(* IEC 61131-3 sources: trust-platform/examples/OSCAT/booster_commissioning_decorator/oop/src, 3 files *)

(* ---- Main.st ---- *)
(* Pattern role: ISignalSource is the contract boundary for the Decorator example. *)
INTERFACE ISignalSource
    PROPERTY Value : REAL
    GET
    END_GET
    END_PROPERTY

    PROPERTY Quality : BYTE
    GET
    END_GET
    END_PROPERTY

    METHOD Update
    END_METHOD
END_INTERFACE

(* Pattern role: IPump is the contract boundary for the Decorator example. *)
INTERFACE IPump
    PROPERTY IsRunning : BOOL
    GET
    END_GET
    END_PROPERTY

    METHOD Run
    VAR_INPUT
        SpeedReference : REAL;
    END_VAR
    END_METHOD

    METHOD Stop
    END_METHOD
END_INTERFACE

(* Pattern role: RealPressureSource is a concrete implementation in the Decorator example. *)
FUNCTION_BLOCK RealPressureSource IMPLEMENTS ISignalSource
VAR
    ValueValue : REAL;
    QualityValue : BYTE := BYTE#2;
END_VAR

METHOD PUBLIC Configure
VAR_INPUT
    PressureBar : REAL;
    QualityCode : BYTE;
END_VAR
ValueValue := PressureBar;
QualityValue := QualityCode;
END_METHOD

METHOD PUBLIC Update
END_METHOD

PUBLIC PROPERTY Value : REAL
GET
    Value := ValueValue;
END_GET
END_PROPERTY

PUBLIC PROPERTY Quality : BYTE
GET
    Quality := QualityValue;
END_GET
END_PROPERTY
END_FUNCTION_BLOCK

(* Pattern role: SimulatedPressureDecorator is a concrete implementation in the Decorator example. *)
FUNCTION_BLOCK SimulatedPressureDecorator IMPLEMENTS ISignalSource
VAR
    RealSourceRef : ISignalSource;
    SineGen : SineSignalGenerator;
    UseSimulationValue : BOOL;
    ValueValue : REAL;
    QualityValue : BYTE;
END_VAR

METHOD PUBLIC Wrap
VAR_INPUT
    RealSource : ISignalSource;
    UseSimulation : BOOL;
END_VAR
RealSourceRef := RealSource;
UseSimulationValue := UseSimulation;
SineGen.Initialize();
SineGen.Configure(Period := T#10s, Amplitude := REAL#0.5, Offset := REAL#4.5, Delay := REAL#0.0);
END_METHOD

METHOD PUBLIC SetSimulation
VAR_INPUT
    Enabled : BOOL;
END_VAR
UseSimulationValue := Enabled;
END_METHOD

METHOD PUBLIC Update
RealSourceRef.Update();
IF UseSimulationValue THEN
    ValueValue := SineGen.Update();
    QualityValue := BYTE#2;
ELSE
    ValueValue := RealSourceRef.Value;
    QualityValue := RealSourceRef.Quality;
END_IF;
END_METHOD

PUBLIC PROPERTY Value : REAL
GET
    Value := ValueValue;
END_GET
END_PROPERTY

PUBLIC PROPERTY Quality : BYTE
GET
    Quality := QualityValue;
END_GET
END_PROPERTY

PUBLIC PROPERTY UsingSimulation : BOOL
GET
    UsingSimulation := UseSimulationValue;
END_GET
END_PROPERTY
END_FUNCTION_BLOCK

(* Pattern role: RealPumpDrive is a concrete implementation in the Decorator example. *)
FUNCTION_BLOCK RealPumpDrive IMPLEMENTS IPump
VAR
    RunningValue : BOOL;
    LastSpeedValue : REAL;
END_VAR

METHOD PUBLIC Run
VAR_INPUT
    SpeedReference : REAL;
END_VAR
LastSpeedValue := SpeedReference;
RunningValue := SpeedReference > REAL#0.0;
END_METHOD

METHOD PUBLIC Stop
LastSpeedValue := REAL#0.0;
RunningValue := FALSE;
END_METHOD

PUBLIC PROPERTY IsRunning : BOOL
GET
    IsRunning := RunningValue;
END_GET
END_PROPERTY

PUBLIC PROPERTY LastSpeed : REAL
GET
    LastSpeed := LastSpeedValue;
END_GET
END_PROPERTY
END_FUNCTION_BLOCK

(* Pattern role: CommissioningOutputDriver is a concrete implementation in the Decorator example. *)
FUNCTION_BLOCK CommissioningOutputDriver IMPLEMENTS IPump
VAR
    RealPump : IPump;
    LoopbackOnlyValue : BOOL;
    LastCommandedSpeedValue : REAL;
END_VAR

METHOD PUBLIC Wrap
VAR_INPUT
    Pump : IPump;
    LoopbackOnly : BOOL;
END_VAR
RealPump := Pump;
LoopbackOnlyValue := LoopbackOnly;
END_METHOD

METHOD PUBLIC SetLoopback
VAR_INPUT
    Enabled : BOOL;
END_VAR
LoopbackOnlyValue := Enabled;
END_METHOD

METHOD PUBLIC Run
VAR_INPUT
    SpeedReference : REAL;
END_VAR
LastCommandedSpeedValue := SpeedReference;
IF NOT LoopbackOnlyValue THEN
    RealPump.Run(SpeedReference := SpeedReference);
END_IF;
END_METHOD

METHOD PUBLIC Stop
LastCommandedSpeedValue := REAL#0.0;
IF NOT LoopbackOnlyValue THEN
    RealPump.Stop();
END_IF;
END_METHOD

PUBLIC PROPERTY IsRunning : BOOL
GET
    IF LoopbackOnlyValue THEN
        IsRunning := LastCommandedSpeedValue > REAL#0.0;
    ELSE
        IsRunning := RealPump.IsRunning;
    END_IF;
END_GET
END_PROPERTY

PUBLIC PROPERTY LastCommandedSpeed : REAL
GET
    LastCommandedSpeed := LastCommandedSpeedValue;
END_GET
END_PROPERTY
END_FUNCTION_BLOCK

(* Composition role: BoosterCommissioningCell owns the collaborating objects used by this Decorator example. *)
FUNCTION_BLOCK BoosterCommissioningCell
VAR
    RealPressure : RealPressureSource;
    PressureDecorator : SimulatedPressureDecorator;
    RealPump : RealPumpDrive;
    PumpDecorator : CommissioningOutputDriver;
    Pressure : ISignalSource;
    Pump : IPump;
END_VAR

METHOD PUBLIC Initialize
RealPressure.Configure(PressureBar := REAL#4.0, QualityCode := BYTE#2);
PressureDecorator.Wrap(RealSource := RealPressure, UseSimulation := FALSE);
PumpDecorator.Wrap(Pump := RealPump, LoopbackOnly := FALSE);
Pressure := PressureDecorator;
Pump := PumpDecorator;
END_METHOD

METHOD PUBLIC Update : REAL
VAR_INPUT
    RealPressureBar : REAL;
    CommissioningMode : BOOL;
    LoopbackOnly : BOOL;
    PressureSetpoint : REAL;
END_VAR
VAR
    SpeedCommand : REAL;
END_VAR
RealPressure.Configure(PressureBar := RealPressureBar, QualityCode := BYTE#2);
PressureDecorator.SetSimulation(Enabled := CommissioningMode);
PumpDecorator.SetLoopback(Enabled := LoopbackOnly);
Pressure.Update();
IF Pressure.Value < PressureSetpoint THEN
    SpeedCommand := REAL#50.0;
    Pump.Run(SpeedReference := SpeedCommand);
ELSE
    Pump.Stop();
END_IF;
Update := SpeedCommand;
END_METHOD

PUBLIC PROPERTY PressureValue : REAL
GET
    PressureValue := Pressure.Value;
END_GET
END_PROPERTY

PUBLIC PROPERTY PressureQuality : BYTE
GET
    PressureQuality := Pressure.Quality;
END_GET
END_PROPERTY

PUBLIC PROPERTY LastCommandedSpeed : REAL
GET
    LastCommandedSpeed := PumpDecorator.LastCommandedSpeed;
END_GET
END_PROPERTY

PUBLIC PROPERTY RealPumpRunning : BOOL
GET
    RealPumpRunning := RealPump.IsRunning;
END_GET
END_PROPERTY
END_FUNCTION_BLOCK

(* Scan role: Main wires the example objects and exposes the PLC call path under test. *)
PROGRAM Main
VAR
    Cell : BoosterCommissioningCell;
    CommissioningMode : BOOL;
    LoopbackOnly : BOOL;
    RealPressureRaw : INT;
    PumpSpeedRaw : INT;
    TestLampOut : BOOL;
END_VAR

Cell.Initialize();
PumpSpeedRaw := REAL_TO_INT(Cell.Update(RealPressureBar := INT_TO_REAL(RealPressureRaw) / REAL#10.0, CommissioningMode := CommissioningMode, LoopbackOnly := LoopbackOnly, PressureSetpoint := REAL#4.5));
TestLampOut := CommissioningMode;
END_PROGRAM

(* ---- Configuration.st ---- *)
CONFIGURATION BoosterCommissioningDecoratorOopConfiguration
RESOURCE Cpu0 ON PLC
    TASK MainTask (INTERVAL := T#100ms, PRIORITY := 1);
    PROGRAM Cell WITH MainTask : Main;
END_RESOURCE
VAR_CONFIG
    Cell.CommissioningMode AT %IX0.0 : BOOL;
    Cell.LoopbackOnly AT %IX0.1 : BOOL;
    Cell.RealPressureRaw AT %IW0 : INT;
    Cell.PumpSpeedRaw AT %QW0 : INT;
    Cell.TestLampOut AT %QX0.0 : BOOL;
END_VAR
END_CONFIGURATION

(* ---- Tests.st ---- *)
TEST_PROGRAM CommissioningPressureDecoratorSubstitutesSimulation
VAR
    Cell : BoosterCommissioningCell;
    Speed : REAL;
END_VAR

Cell.Initialize();
Speed := Cell.Update(RealPressureBar := REAL#9.0, CommissioningMode := TRUE, LoopbackOnly := TRUE, PressureSetpoint := REAL#4.5);
ASSERT_EQUAL(EXPECTED := BYTE#2, ACTUAL := Cell.PressureQuality);
ASSERT_TRUE(IN := Cell.LastCommandedSpeed >= REAL#0.0);
ASSERT_FALSE(IN := Cell.RealPumpRunning);
END_TEST_PROGRAM

TEST_PROGRAM CommissioningOutputDriverLoopbackDoesNotRunRealPump
VAR
    RealPump : RealPumpDrive;
    Wrapper : CommissioningOutputDriver;
END_VAR

Wrapper.Wrap(Pump := RealPump, LoopbackOnly := TRUE);
Wrapper.Run(SpeedReference := REAL#60.0);
ASSERT_NEAR(EXPECTED := REAL#60.0, ACTUAL := Wrapper.LastCommandedSpeed, DELTA := REAL#0.001);
ASSERT_FALSE(IN := RealPump.IsRunning);
ASSERT_TRUE(IN := Wrapper.IsRunning);
END_TEST_PROGRAM

(* Mode-switch test: same cell instance runs in commissioning mode then
   in production mode. Catches bugs where the decorator caches its
   wrapped state from a previous mode, or where switching from loopback
   to live unintentionally leaves the real pump running from earlier
   simulated commands. *)
TEST_PROGRAM CommissioningCellSwitchesBetweenSimAndLiveOnSameInstance
VAR
    Cell : BoosterCommissioningCell;
    SimSpeed : REAL;
    LiveSpeed : REAL;
END_VAR

Cell.Initialize();

(* Scan 1: commissioning + loopback -> simulated path, no real pump *)
SimSpeed := Cell.Update(RealPressureBar := REAL#9.0, CommissioningMode := TRUE, LoopbackOnly := TRUE, PressureSetpoint := REAL#4.5);
ASSERT_FALSE(IN := Cell.RealPumpRunning);

(* Scan 2: production mode (live signal, live pump) on same instance *)
LiveSpeed := Cell.Update(RealPressureBar := REAL#3.0, CommissioningMode := FALSE, LoopbackOnly := FALSE, PressureSetpoint := REAL#4.5);
(* Quality must reflect the live source, not the previous sim quality *)
ASSERT_EQUAL(EXPECTED := BYTE#2, ACTUAL := Cell.PressureQuality);
END_TEST_PROGRAM

(* RealPressureSource isolation: returns configured value/quality. *)
TEST_PROGRAM RealPressureSourceReturnsConfiguredValue
VAR
    Source : RealPressureSource;
END_VAR
Source.Configure(PressureBar := REAL#7.5, QualityCode := BYTE#1);
Source.Update();
ASSERT_NEAR(EXPECTED := REAL#7.5, ACTUAL := Source.Value, DELTA := REAL#0.001);
ASSERT_EQUAL(EXPECTED := BYTE#1, ACTUAL := Source.Quality);

(* Reconfigure: new values reflected after next read *)
Source.Configure(PressureBar := REAL#3.2, QualityCode := BYTE#0);
Source.Update();
ASSERT_NEAR(EXPECTED := REAL#3.2, ACTUAL := Source.Value, DELTA := REAL#0.001);
ASSERT_EQUAL(EXPECTED := BYTE#0, ACTUAL := Source.Quality);
END_TEST_PROGRAM

(* SimulatedPressureDecorator forwards real source when simulation is off. *)
TEST_PROGRAM SimulatedPressureDecoratorForwardsRealWhenSimOff
VAR
    LiveSource : RealPressureSource;
    Decorator : SimulatedPressureDecorator;
END_VAR
LiveSource.Configure(PressureBar := REAL#5.5, QualityCode := BYTE#2);
Decorator.Wrap(RealSource := LiveSource, UseSimulation := FALSE);
Decorator.Update();
ASSERT_NEAR(EXPECTED := REAL#5.5, ACTUAL := Decorator.Value, DELTA := REAL#0.001);
ASSERT_FALSE(IN := Decorator.UsingSimulation);

(* Switch to simulation: value comes from sine generator, not real *)
Decorator.SetSimulation(Enabled := TRUE);
Decorator.Update();
ASSERT_TRUE(IN := Decorator.UsingSimulation);
END_TEST_PROGRAM

(* RealPumpDrive isolation: Run sets running, Stop clears it. *)
TEST_PROGRAM RealPumpDriveTracksRunStop
VAR
    Pump : RealPumpDrive;
END_VAR
ASSERT_FALSE(IN := Pump.IsRunning);
Pump.Run(SpeedReference := REAL#42.0);
ASSERT_TRUE(IN := Pump.IsRunning);
ASSERT_NEAR(EXPECTED := REAL#42.0, ACTUAL := Pump.LastSpeed, DELTA := REAL#0.001);

Pump.Stop();
ASSERT_FALSE(IN := Pump.IsRunning);
ASSERT_NEAR(EXPECTED := REAL#0.0, ACTUAL := Pump.LastSpeed, DELTA := REAL#0.001);

(* Run with zero speed should not flag running *)
Pump.Run(SpeedReference := REAL#0.0);
ASSERT_FALSE(IN := Pump.IsRunning);
END_TEST_PROGRAM

(* Cell control loop: pressure below setpoint runs pump, above stops. *)
TEST_PROGRAM CommissioningCellControlBoundary
VAR
    Cell : BoosterCommissioningCell;
END_VAR
Cell.Initialize();

(* Below setpoint: pump runs *)
Cell.Update(RealPressureBar := REAL#3.0, CommissioningMode := FALSE, LoopbackOnly := FALSE, PressureSetpoint := REAL#4.5);
ASSERT_TRUE(IN := Cell.RealPumpRunning);

(* At setpoint: pump stops (strict inequality) *)
Cell.Update(RealPressureBar := REAL#4.5, CommissioningMode := FALSE, LoopbackOnly := FALSE, PressureSetpoint := REAL#4.5);
ASSERT_FALSE(IN := Cell.RealPumpRunning);

(* Above setpoint: pump stops *)
Cell.Update(RealPressureBar := REAL#5.0, CommissioningMode := FALSE, LoopbackOnly := FALSE, PressureSetpoint := REAL#4.5);
ASSERT_FALSE(IN := Cell.RealPumpRunning);
END_TEST_PROGRAM
